(* IEC 61131-3 sources: s7-to-codesys/tests/POUs/Graph/FB_BackwashGraph_SeqTest, 11 files *)

(* ---- FB_BackwashGraph_SeqTest.decl.st ---- *)
// Назначение: многоцикловый набор CfUnit (coUnit 1.2.0.0) без времени для FB_BackwashGraph — промывки
//             фильтра, переведённой из S7-GRAPH. Один и тот же набор проходят оба варианта: ST-двойник
//             (src/POUs/Lang/Converted, этот проект) и SFC с ФБ-обёрткой (plcopen/Lang/Converted, проект
//             tools_project/cds_plcopen.py test). SFC переключается в конце цикла, двойник — в том же вызове,
//             поэтому каждый шаг теста — CYCLES вызовов с одинаковыми входами, затем проверки установившегося
//             состояния. Пути с временем (продувка 10 с, D задвижки воздуха) проверяют сценарии ST-двойника.
//             Ожидаемые значения — по описанию блока (samples/lang/README.md), а не по результату перевода.
//             Экземпляр набора объявляется в PRG_Tests.
// Автор:      kr0nsch
// Версия:     1.2.0
// Документ:   docs/MAPPING_GRAPH.md; docs/EQUIVALENCE.md
FUNCTION_BLOCK FB_BackwashGraph_SeqTest EXTENDS coUnit.FB_TestSuite
VAR CONSTANT
    CYCLES : INT := 3;  // вызовов на шаг теста: хватает SFC (переключение в конце цикла) и двойнику
END_VAR

(* ---- InitResets.method.decl.st ---- *)
// INIT_SQ возвращает начальный шаг (действия Drain выключены) и держит его; после снятия — новый пуск,
// промывка №2 (событие S1 — один раз).
METHOD PRIVATE InitResets
VAR
    fbDut : FB_BackwashGraph;   // проверяемый блок
    iCycle : INT;               // вызов внутри шага теста
END_VAR

(* ---- InitResets.method.impl.st ---- *)
coUnit.TEST('InitResets');
FOR iCycle := 1 TO CYCLES DO
    fbDut(xStart := TRUE);
END_FOR
AssertTrue(Condition := fbDut.xDrainValve, Message := 'Drain');

FOR iCycle := 1 TO CYCLES DO
    fbDut(INIT_SQ := TRUE);
END_FOR
AssertTrue(Condition := fbDut.xReady, Message := 'INIT_SQ: Idle');
AssertFalse(Condition := fbDut.xDrainValve, Message := 'INIT_SQ: drain closed');

FOR iCycle := 1 TO CYCLES DO
    fbDut(INIT_SQ := FALSE, xStart := TRUE);
END_FOR
AssertTrue(Condition := fbDut.xDrainValve, Message := 'restart: Drain');
AssertEquals_INT(Expected := 2, Actual := fbDut.iWashCount, Message := 'wash #2');
coUnit.TEST_FINISHED();

(* ---- InterlockStopsPump.method.decl.st ---- *)
// Блокировка шага Rinse (NC): при неисправном насосе (xPumpOk = FALSE) насос промывки выключен, воздуходувка
// параллельного шага работает; насос исправен — снова включён.
METHOD PRIVATE InterlockStopsPump
VAR
    fbDut : FB_BackwashGraph;   // проверяемый блок
    iCycle : INT;               // вызов внутри шага теста
END_VAR

(* ---- InterlockStopsPump.method.impl.st ---- *)
coUnit.TEST('InterlockStopsPump');
FOR iCycle := 1 TO CYCLES DO
    fbDut(xStart := TRUE);
END_FOR
FOR iCycle := 1 TO CYCLES DO
    fbDut(xStart := FALSE, xLevelLow := TRUE);
END_FOR
AssertTrue(Condition := fbDut.xWashPump, Message := 'Rinse: pump');

FOR iCycle := 1 TO CYCLES DO
    fbDut(xLevelLow := FALSE, xPumpOk := FALSE);
END_FOR
AssertFalse(Condition := fbDut.xWashPump, Message := 'interlock not met: pump off');
AssertTrue(Condition := fbDut.xBlower, Message := 'Air keeps running');

FOR iCycle := 1 TO CYCLES DO
    fbDut(xPumpOk := TRUE);
END_FOR
AssertTrue(Condition := fbDut.xWashPump, Message := 'interlock met: pump on');
coUnit.TEST_FINISHED();

(* ---- LongWashParallel.method.decl.st ---- *)
// Длинная промывка: после слива параллельно Air (воздуходувка) и Rinse (насос); задвижка воздуха (D 2 с) без
// времени закрыта.
METHOD PRIVATE LongWashParallel
VAR
    fbDut : FB_BackwashGraph;   // проверяемый блок
    iCycle : INT;               // вызов внутри шага теста
END_VAR

(* ---- LongWashParallel.method.impl.st ---- *)
coUnit.TEST('LongWashParallel');
FOR iCycle := 1 TO CYCLES DO
    fbDut(xStart := TRUE);
END_FOR
AssertTrue(Condition := fbDut.xDrainValve, Message := 'Drain');

FOR iCycle := 1 TO CYCLES DO
    fbDut(xStart := FALSE, xLevelLow := TRUE);
END_FOR
AssertFalse(Condition := fbDut.xDrainValve, Message := 'parallel: drain closed');
AssertTrue(Condition := fbDut.xBlower, Message := 'parallel: Air blower');
AssertTrue(Condition := fbDut.xWashPump, Message := 'parallel: Rinse pump');
AssertFalse(Condition := fbDut.xAirValve, Message := 'D 2 s not elapsed');
AssertTrue(Condition := fbDut.xWashActive, Message := 'wash active');
coUnit.TEST_FINISHED();

(* ---- ShortWashCycle.method.decl.st ---- *)
// Короткая промывка целиком: Idle → Drain (S1: промывка №1) → QuickRinse → Refill → Idle.
METHOD PRIVATE ShortWashCycle
VAR
    fbDut : FB_BackwashGraph;   // проверяемый блок (новый экземпляр на каждый вызов метода)
    iCycle : INT;               // вызов внутри шага теста
END_VAR

(* ---- ShortWashCycle.method.impl.st ---- *)
coUnit.TEST('ShortWashCycle');
FOR iCycle := 1 TO CYCLES DO
    fbDut();
END_FOR
AssertTrue(Condition := fbDut.xReady, Message := 'Idle: ready');
AssertFalse(Condition := fbDut.xDrainValve, Message := 'Idle: drain closed');

FOR iCycle := 1 TO CYCLES DO
    fbDut(xStart := TRUE);
END_FOR
AssertFalse(Condition := fbDut.xReady, Message := 'Drain: not ready');
AssertTrue(Condition := fbDut.xDrainValve, Message := 'Drain: drain open');
AssertTrue(Condition := fbDut.xWashActive, Message := 'Drain: S wash active');
AssertTrue(Condition := fbDut.xValvesBusy, Message := 'Drain: post operation');
AssertEquals_INT(Expected := 1, Actual := fbDut.iWashCount, Message := 'Drain: S1 count once');

FOR iCycle := 1 TO CYCLES DO
    fbDut(xStart := FALSE, xLevelLow := TRUE, xShortWash := TRUE);
END_FOR
AssertFalse(Condition := fbDut.xDrainValve, Message := 'QuickRinse: drain closed');
AssertTrue(Condition := fbDut.xWashPump, Message := 'QuickRinse: pump');
AssertFalse(Condition := fbDut.xBlower, Message := 'QuickRinse: no blower');

FOR iCycle := 1 TO CYCLES DO
    fbDut(xLevelLow := FALSE, xLevelHigh := TRUE);
END_FOR
AssertTrue(Condition := fbDut.xReady, Message := 'back to Idle');
AssertFalse(Condition := fbDut.xWashPump, Message := 'Idle: pump off');
AssertFalse(Condition := fbDut.xInletValve, Message := 'Idle: inlet closed');
AssertFalse(Condition := fbDut.xWashActive, Message := 'Refill: R wash active');
AssertEquals_INT(Expected := 1, Actual := fbDut.iWashCount, Message := 'one wash');
coUnit.TEST_FINISHED();

(* ---- SupervisionHoldsUntilAck.method.decl.st ---- *)
// Контроль шага Drain: неисправность задвижки защёлкивает ошибку (ERR_FLT), переход заблокирован и после
// ухода неисправности; квитирование ACK_EF снимает ошибку, и переход проходит.
METHOD PRIVATE SupervisionHoldsUntilAck
VAR
    fbDut : FB_BackwashGraph;   // проверяемый блок
    iCycle : INT;               // вызов внутри шага теста
END_VAR

(* ---- SupervisionHoldsUntilAck.method.impl.st ---- *)
coUnit.TEST('SupervisionHoldsUntilAck');
FOR iCycle := 1 TO CYCLES DO
    fbDut(xStart := TRUE);
END_FOR
FOR iCycle := 1 TO CYCLES DO
    fbDut(xStart := FALSE, xValveFault := TRUE);
END_FOR
AssertTrue(Condition := fbDut.ERR_FLT, Message := 'supervision error');

FOR iCycle := 1 TO CYCLES DO
    fbDut(xValveFault := FALSE, xLevelLow := TRUE, xShortWash := TRUE);
END_FOR
AssertTrue(Condition := fbDut.ERR_FLT, Message := 'error latched');
AssertTrue(Condition := fbDut.xDrainValve, Message := 'transition blocked: still Drain');
AssertFalse(Condition := fbDut.xWashPump, Message := 'no QuickRinse yet');

FOR iCycle := 1 TO CYCLES DO
    fbDut(ACK_EF := TRUE);
END_FOR
AssertFalse(Condition := fbDut.ERR_FLT, Message := 'acknowledged');
AssertFalse(Condition := fbDut.xDrainValve, Message := 'Drain left');
AssertTrue(Condition := fbDut.xWashPump, Message := 'QuickRinse');
coUnit.TEST_FINISHED();
